Universal Robots URScript: T012_codellama_34b_adversarial_A8.4_rep1.urscript

def program():
    # Home the robot
    movej(p[0, 0, 0, 0, 0, 0], v=200.0)

    # Approach spot 1
    movel(p[0, 0, 0, 0, 0, -200], v=200.0)

    # Descend
